# EPICS autosave request: iocs/ad/simdetector-ioc/auto_settings.req
file "simDetector_settings.req",    P=$(P),  R=cam1:
file "NDStdArrays_settings.req",    P=$(P),  R=image1:
file "NDStdArrays_settings.req",    P=$(P),  R=image2:
file "commonPlugin_settings.req",   P=$(P)
